// TIA Portal V20 export
// export: Created 2026-10-19T18:04:31.5918765Z, ExportSetting WithDefaults, DisplayName Totally Integrated Automation Portal, DisplayVersion V20 Update 6, DisplayName TIA Portal Openness, DisplayVersion V20 Update 6, DisplayName TIA Portal Version Control Interface, DisplayVersion V20 Update 6, DisplayName SINAMICS Startdrive Advanced, DisplayVersion V20 SP1, DisplayName SINAMICS Startdrive G130, G150, S120, S150, SINAMICS MV, G220, S200, S210, DisplayVersion V20 SP1, DisplayName SINAMICS Startdrive G110M, G120, G120C, G120D, G120P, G115D, DisplayVersion V20 SP1, DisplayName STEP 7 Professional, DisplayVersion V20 Update 6, DisplayName STEP 7 Safety, DisplayVersion V20 Update 2, DisplayName WinCC Basic/Comfort/Advanced, DisplayVersion V20 Update 6, DisplayName WinCC Unified, DisplayVersion V20 Update 6
DATA_BLOCK "Screen_DB"   // DB23
{ S7_Optimized_Access := 'TRUE' }
VERSION : 0.1
// stored: AutoNumber true, DBAccessibleFromOPCUA true, DBAccessibleFromWebserver true, IsOnlyStoredInLoadMemory false, IsRetainMemResEnabled false, IsWriteProtectedInAS false, MemoryReserve 100
   VAR
      VTD_LevelDetect { S7_SetPoint := 'True'} : Array[1..8] of Bool;
      VTD_Semi_CMD : Array[1..8] of Bool;
      VTD_ActualPosition { S7_SetPoint := 'True'} : DInt;
      VTD_OvertravelUp : Bool;
      VTD_LimitUp : Bool;
      VTD_CreepUp : Bool;
      VTD_SlowDownUp : Bool;
      VTD_SlowDownDown : Bool;
      VTD_CreepDown : Bool;
      VTD_LimitDown : Bool;
      VTD_OvertravelDown : Bool;
      VTD_LiftUp : Bool;
      VTD_LiftDown : Bool;
      VTD_LimitOverride : Bool;
      VTD_Manual : Bool;
      VTD_Semi : Bool;
      VTD_MemoryLatch : Bool;
      VTD_SaveData : Bool;
      VTD_Select : USInt;
      Cnv_Manual : Bool;
      Cnv_Semi : Bool;
      Cnv_Foward : Bool;
      Cnv_Backward : Bool;
      Cnv_LeftAllign : Bool;
      Cnv_RightAllign : Bool;
      Cnv_FowardTransfer : Bool;
      Cnv_BackwardTransfer : Bool;
      Cnv_ShuttleStopper : Bool;
      Cnv_ShuttleStopperVisibility : Bool;
      Cnv_Plallet_Type1Visibility : Bool;
      Cnv_Plallet_Type2Visibility : Bool;
      Cnv_Select : USInt;
      Shuttle_Status : "Shuttle_MQTT_Status_Msg";
      Shuttle_Name { S7_SetPoint := 'True'} : String;
      Shuttle_URL : String;
      Settings_ActivePopUp : USInt;
      Alarms_ActiveTable : USInt;
      MainTemplate_ErrorActive : Bool;
      MainTemplate_ErrorCount : USInt;
      MainTemplate_ScreenNo : UInt;
      MainTemplate_Background : USInt;
      EmptyTemplate_Background : USInt;
      IO_ActivePopup : USInt;
      Charge_VTD : Bool;
      Charge_Cnv : Bool;
      Charge_VTD_Commands : Bool;
      Charge_Cnv_Commands : Bool;
      Shuttle : "Shuttle_MQTT_Status_Msg";
      Shuttle_Select : USInt;
   END_VAR
BEGIN
END_DATA_BLOCK
